(*
SPDX-FileCopyrightText: c 2026 Oleksandr Tiutyk <trofimich@gmail.com>
SPDX-License-Identifier: MIT
License: https://opensource.org/license/mit
*)

(*!
<summary>Groups byte-string builder assignment, reuse and failure contracts.</summary>
<description>
Owns the independent child instances and their fixed registration array. Use from one PLC task at a stable address.
</description>
*)

{attribute 'no_assign'}
{attribute 'no_explicit_call' := 'do not call this function block directly'}
FUNCTION_BLOCK StringBuilderTestGroup EXTENDS TOF_Testing.TestGroup<3>
VAR_STAT
	{attribute 'hide'}
	_ClassName : STRING := __POUNAME();
END_VAR
VAR
	_BuildEmpty : StringBuilderEmptyTest(name := "BuildEmpty", parent := THIS^);
	_BuildNotEmpty : StringBuilderContentTest(name := "BuildNotEmpty", parent := THIS^);
	_ErrorChecking : StringBuilderAssignmentFailureTest(name := "ErrorChecking", parent := THIS^);

	_Children : ARRAY [0.._ChildCount - 1] OF TOF_Testing.ITestElement :=
	[
		_BuildEmpty,
		_BuildNotEmpty,
		_ErrorChecking
	];
END_VAR

//! <summary>Borrows the fixed child array. Callers must not modify it.</summary>
{attribute 'monitoring' := 'call'}
PROPERTY Children : REFERENCE TO ARRAY [0.._ChildCount - 1] OF TOF_Testing.ITestElement
GET
Children REF= _Children;
END_GET
END_PROPERTY

//! <summary>Borrows the concrete class name. Callers must not modify it.</summary>
{attribute 'monitoring' := 'call'}
PROPERTY ClassName : REFERENCE TO STRING
GET
ClassName REF= _ClassName;
END_GET
END_PROPERTY

//! <summary>Borrows the compiler-initialized namespace name. Callers must not modify it.</summary>
{attribute 'monitoring' := 'call'}
PROPERTY NamespaceName : REFERENCE TO STRING
GET
NamespaceName REF= CurrentNamespace.Name;
END_GET
END_PROPERTY

//! <summary>Reports the concrete instance size in bytes.</summary>
{attribute 'monitoring' := 'call'}
PROPERTY SelfSize : ULINT
GET
SelfSize := XSIZEOF(THIS^);
END_GET
END_PROPERTY

END_FUNCTION_BLOCK

(* stored: Version 1.1.0.1
   POU StringBuilderTestGroup: Id {0ff202ab-ff5f-47eb-bea4-d472be3897c7}, SpecialFunc None
   Property Children: Id {57c0c710-87ec-46d2-bf82-cf780307d09f}
   Get Get: Id {a573e352-0f07-4a3c-b8e6-8c13da48b43d}
   Property ClassName: Id {48e632ce-16c4-4aaa-9822-7cfdf34ec3ec}
   Get Get: Id {8bee5897-75d5-42e5-a331-129b6de09cce}
   Property NamespaceName: Id {44ecaa0f-f3c3-4f8e-a1e1-fdf3690a49df}
   Get Get: Id {37e630d0-6a2c-4280-adc2-92dbfa333110}
   Property SelfSize: Id {3a91a2b9-6188-46c5-ae29-a46b782c2cba}
   Get Get: Id {7e5972fb-2c76-4be3-92e4-9ff539761160} *)
